// TIA Portal V19 export
TYPE "ST_PICK_POSITION"
   STRUCT
      Pick : Array[0..50] of "ST_Pos";
      iLastPick { S7_SetPoint := 'True'} : Int;
   END_STRUCT;
END_TYPE
